(* PLC project , Example Fixture *)

FUNCTION F_Acc : INT
  VAR_INPUT
    n : INT;
  END_VAR
  VAR
    acc : INT;
  END_VAR

IF acc > n THEN (* PLCA-Q010 *)
    F_Acc := 1;
END_IF
acc := n;
END_FUNCTION
